PROGRAM MAIN
VAR
    fbCamMachine : FB_CamMachine;
END_VAR

fbCamMachine(
    stCommands := GVL_CamControl.stCommands,
    stRecipe := GVL_CamControl.stRecipe,
    AxisConveyor := GVL_Motion.gAxisConveyor,
    AxisCutter := GVL_Motion.gAxisCutter,
    stStatus => GVL_CamControl.stStatus,
    stScope => GVL_CamControl.stScope);

END_PROGRAM

(* stored: Version 1.1.0.1, ProductVersion 3.1.4024.16
   POU MAIN: Id {4a4be6dc-9e2b-467b-a657-9d8f59dc44c0}, SpecialFunc None *)
